TYPE ST_DataHistoryHMI :
STRUCT
    iNestIndex 		: INT;
    sResult 		: STRING(10);
    rDistance  		: REAL;
    rForce     		: REAL;
    dtTimeStamp 	: DATE_AND_TIME;
END_STRUCT
END_TYPE

(* stored: Version 1.1.0.1
   DUT ST_DataHistoryHMI: Id {6478a192-85c4-42dd-85bd-7d4a007ddc4a} *)
